(* IEC 61131-3 sources: kns-port-domestic/upstream/kns-pump-station/src/DUTs/Station, 10 files *)

(* ---- E_ControlAct.dut.st ---- *)
// Назначение: действующее управление насосами (04 §4), поле stStationSts.eControlAct.
//             Старшинство в «Автомате»: PowerLost > Restart > DryRunStop > Float > Emergency >
//             LevelPid > Stepped.
// Автор:      kr0nsch
// Версия:     0.1.0
// Документ:   docs/DESIGN.md, раздел 3.1
{attribute 'qualified_only'}
{attribute 'strict'}
TYPE E_ControlAct :
(
    Manual     := 0,   // станция в «Ручном»: запросов нет, только блокировки
    Stepped    := 1,   // ступенчатое регулирование
    LevelPid   := 2,   // ПИД уровня и подключение по нагрузке
    Float      := 3,   // резервное управление по поплавкам (LT101 недостоверен)
    Emergency  := 4,   // аварийно высокий уровень: все доступные насосы
    DryRunStop := 5,   // защита «сухой ход»: запросы сняты
    PowerLost  := 6,   // нет напряжения на вводе
    Restart    := 7    // задержка после старта или восстановления питания, последовательный пуск
) INT;
END_TYPE

(* ---- E_ControlMethod.dut.st ---- *)
// Назначение: выбранный способ регулирования (04 §3.2, 18.2 № 1). Другое значение в retain
//             санитизируется в Stepped.
// Автор:      kr0nsch
// Версия:     0.1.0
// Документ:   docs/DESIGN.md, раздел 3.1
{attribute 'qualified_only'}
{attribute 'strict'}
TYPE E_ControlMethod :
(
    Stepped  := 1,   // ступенчатое по уровням (04 §6)
    LevelPid := 2    // поддержание уровня ПИД LIC101 (04 §7)
) INT;
END_TYPE

(* ---- E_PumpRole.dut.st ---- *)
// Назначение: роль насоса в станции (04 §5.1).
// Автор:      kr0nsch
// Версия:     0.1.0
// Документ:   docs/DESIGN.md, раздел 3.1
{attribute 'qualified_only'}
{attribute 'strict'}
TYPE E_PumpRole :
(
    None    := 0,   // недоступен автоматике (отказ, блокировка, не Auto, нет напряжения)
    Lead    := 1,   // ведущий: запускается первым, в ПИД его частоту регулирует LIC101
    Assist  := 2,   // подпорный: подключается при нехватке производительности
    Standby := 3    // резервный: доступен, не запрошен
) INT;
END_TYPE

(* ---- E_RotationMode.dut.st ---- *)
// Назначение: режим чередования насосов (04 §8.1, 18.2 № 14).
// Автор:      kr0nsch
// Версия:     0.1.0
// Документ:   docs/DESIGN.md, раздел 3.1
{attribute 'qualified_only'}
{attribute 'strict'}
TYPE E_RotationMode :
(
    RunHours := 1,   // по моточасам: меньше RunSeconds, затем меньше Starts, затем меньший номер
    Cyclic   := 2,   // по кругу: следующий после stStationRetain.uiNextLead
    Fixed    := 3    // без чередования: Н1, Н2, Н3
) INT;
END_TYPE

(* ---- E_StationAlarm.dut.st ---- *)
// Назначение: слоты тревог станции KNS1.* (04 §15, 05_alarm_list.csv): индекс массивов
//             FB_StationAlarms и ST_StationCfg.astAlarm; номер тревоги = STN_ALARM_ID_BASE + slot,
//             бит слов wAlm* — slot - 1. Без strict: перечислением индексируются массивы.
// Автор:      kr0nsch
// Версия:     0.1.0
// Документ:   docs/DESIGN.md, раздел 3.1
{attribute 'qualified_only'}
TYPE E_StationAlarm :
(
    EHL    := 1,    // аварийно высокий уровень (Critical)
    DRY    := 2,    // сухой ход станции (High)
    LACK   := 3,    // недостаточно насосов (High)
    NORES  := 4,    // нет резерва (High)
    ATS    := 5,    // АВР выполнен (Medium)
    FLOAT  := 6,    // управление по поплавкам (Medium)
    LDEV   := 7,    // противоречие поплавка и уровнемера (Medium)
    STEP   := 8,    // ступенчатое вместо ПИД (Low)
    NOAUTO := 9,    // станция в «Ручном» дольше 600 с (Low)
    UL1    := 10,   // недогрузка (сухой ход) Н1 (Medium)
    UL2    := 11,   // недогрузка Н2
    UL3    := 12,   // недогрузка Н3
    SIM    := 13    // режим имитации (Low)
) UINT;
END_TYPE

(* ---- E_StationMode.dut.st ---- *)
// Назначение: режим станции (04 §3). Другое значение в retain санитизируется в Manual
//             сравнениями (FB_StationMode, правило L4 контракта plc-process-lib).
// Автор:      kr0nsch
// Версия:     0.1.0
// Документ:   docs/DESIGN.md, раздел 3.1
{attribute 'qualified_only'}
{attribute 'strict'}
TYPE E_StationMode :
(
    Auto   := 1,   // «Автомат»: насосами управляет логика станции
    Manual := 2    // «Ручной»: насосами управляет оператор с HMI, блокировки действуют
) INT;
END_TYPE

(* ---- ST_StationCfg.dut.st ---- *)
// Назначение: уставки станции (GVL_Persist.stStationCfg) — параметры 04 §18.2 № 2–31 с теми же
//             именами и значениями по умолчанию, тревоги KNS1.* и резерв. Значения по умолчанию
//             проходят F_StationCfgCheck. Тип лежит в Persistent Variables и заморожен целиком:
//             новые параметры 1.x — в элементах резерва без переименования.
// Автор:      kr0nsch
// Версия:     0.1.0
// Документ:   docs/DESIGN.md, раздел 3.1
{attribute 'qualified_only'}
TYPE ST_StationCfg :
STRUCT
    // уровни (№ 2–6)
    rLvlStop_m          : REAL := 1.00;
    rLvlStartLead_m     : REAL := 1.60;
    rLvlStopAssist_m    : REAL := 1.40;
    rLvlStartAssist_m   : REAL := 2.40;
    tLvlConfirm         : TIME := T#5S;
    // ступенчатое (№ 7)
    rStepSpeed_pct      : REAL := 100.0;
    // ПИД (№ 8–12)
    rLevelSp_m          : REAL := 1.40;
    rAssistOn_pct       : REAL := 98.0;
    tAssistOn           : TIME := T#30S;
    rAssistOff_pct      : REAL := 75.0;
    tAssistOff          : TIME := T#60S;
    // роли (№ 13–17)
    uiDutyMax           : UINT := 2;
    eRotation           : E_RotationMode := E_RotationMode.RunHours;
    tMaxContRun         : TIME := T#4H;
    tOverlap            : TIME := T#10S;
    tStagger            : TIME := T#5S;
    // питание (№ 18–20)
    tPwrRestart         : TIME := T#10S;
    tSeqStep            : TIME := T#15S;
    tPlcStart           : TIME := T#10S;
    // защиты (№ 21–27)
    tDryRelease         : TIME := T#60S;
    rLdev102On_m        : REAL := 3.50;
    rLdev102Off_m       : REAL := 4.40;
    rLdev103On_m        : REAL := 0.80;
    rLdev103Off_m       : REAL := 0.20;
    tLdev               : TIME := T#30S;
    tLtRecover          : TIME := T#30S;
    // недогрузка (№ 28–30)
    rUnderload_A        : REAL := 12.0;
    rUnderloadSpeed_pct : REAL := 80.0;
    tUnderload          : TIME := T#15S;
    // вентиляция (№ 31)
    tV1Overrun          : TIME := T#10M;
    // тревоги KNS1.* по 05_alarm_list.csv (source = station), индекс — E_StationAlarm. Задержка появления
    // в 05 = tOnDelay + выдержка логики (LDEV — tLdev, UL1…UL3 — tUnderload). Инициализатор — весь
    // массив целиком (правило 3 API 18.3)
    astAlarm            : ARRAY[1..GVL_Const.STN_ALARM_COUNT] OF PL.ST_AlarmCfg := [
        (ePriority := PL.E_AlarmPriority.Critical, tShelveMax := T#0S),   // 1 EHL: откладывать нельзя
        (ePriority := PL.E_AlarmPriority.High),                          // 2 DRY
        (ePriority := PL.E_AlarmPriority.High, tOnDelay := T#10S),       // 3 LACK
        (ePriority := PL.E_AlarmPriority.High, tOnDelay := T#10S),       // 4 NORES
        (ePriority := PL.E_AlarmPriority.Medium),                        // 5 ATS
        (ePriority := PL.E_AlarmPriority.Medium),                        // 6 FLOAT
        (ePriority := PL.E_AlarmPriority.Medium),                        // 7 LDEV
        (ePriority := PL.E_AlarmPriority.Low, tOnDelay := T#10S),        // 8 STEP: без переходных циклов старта
        (ePriority := PL.E_AlarmPriority.Low, tOnDelay := T#10M),        // 9 NOAUTO
        (ePriority := PL.E_AlarmPriority.Medium),                        // 10 UL1
        (ePriority := PL.E_AlarmPriority.Medium),                        // 11 UL2
        (ePriority := PL.E_AlarmPriority.Medium),                        // 12 UL3
        (ePriority := PL.E_AlarmPriority.Low)];                          // 13 SIM
    // резерв: новые параметры 1.x без смены типа; смысл элемента записывается в DESIGN, раздел 3.1
    arReserve           : ARRAY[0..7] OF REAL;
    atReserve           : ARRAY[0..3] OF TIME;
    auiReserve          : ARRAY[0..3] OF UINT;
END_STRUCT
END_TYPE

(* ---- ST_StationCmd.dut.st ---- *)
// Назначение: команды станции (GVL_Station.stStationCmd) — пишут HMI, OPC UA, MQTT. Импульсы и
//             номера обрабатывает и сбрасывает PRG_Station в том же цикле (04 §19.2); результат —
//             stStationSts.eCmdResult и uiCmdSeq.
// Автор:      kr0nsch
// Версия:     0.1.0
// Документ:   docs/DESIGN.md, раздел 3.1
{attribute 'qualified_only'}
TYPE ST_StationCmd :
STRUCT
    xSetAuto      : BOOL;           // импульс: станция в «Автомат» (04 §19.2)
    xSetManual    : BOOL;           // импульс: в «Ручной»; старше xSetAuto
    xSetStepped   : BOOL;           // импульс: способ «ступенчатое»; старше xSetLevelPid
    xSetLevelPid  : BOOL;           // импульс: способ «ПИД уровня»
    xAckAll       : BOOL;           // импульс: квитировать все тревоги станции, LIC101 и устройств
    xResetAll     : BOOL;           // импульс: общий сброс (как HS501)
    xSilence      : BOOL;           // импульс: выключить сирену (как HS502)
    xExportLog    : BOOL;           // импульс: выгрузить журнал в CSV (04 §19.2)
    xRevertCfg    : BOOL;           // импульс: откатить записанные уставки к действующей копии (08 §14, вопрос 2)
    wAckReq       : WORD;           // маска: квитировать тревоги станции, бит slot - 1
    wShelveReq    : WORD;           // маска: отложить на astAlarm[slot].tShelveMax
    wUnshelveReq  : WORD;           // маска: вернуть отложенные
    udiAckId      : UDINT;          // квитировать тревогу по номеру (таблица HMI); 0 — нет; сбрасывается в 0
    udiShelveId   : UDINT;          // отложить тревогу любого источника на её tShelveMax; 0 — нет (08 §14, вопрос 1)
    udiUnshelveId : UDINT;          // вернуть отложенную тревогу по номеру; 0 — нет
END_STRUCT
END_TYPE

(* ---- ST_StationRetain.dut.st ---- *)
// Назначение: энергонезависимое состояние станции (GVL_Persist.stStationRetain): режим, способ
//             регулирования, следующий ведущий для чередования по кругу. Тип лежит в Persistent
//             Variables: не менять (новые данные — в резерве).
// Автор:      kr0nsch
// Версия:     0.1.0
// Документ:   docs/DESIGN.md, раздел 3.1
{attribute 'qualified_only'}
TYPE ST_StationRetain :
STRUCT
    eMode       : E_StationMode := E_StationMode.Manual;      // пустой retain — «Ручной» (04 §3.2)
    eMethod     : E_ControlMethod := E_ControlMethod.Stepped;
    uiNextLead  : UINT := 1;                                  // Cyclic: следующий ведущий
    uiReserve   : UINT;
    audiReserve : ARRAY[0..7] OF UDINT;
END_STRUCT
END_TYPE

(* ---- ST_StationSts.dut.st ---- *)
// Назначение: состояние станции (GVL_Station.stStationSts) для HMI, OPC UA и MQTT: только 16- и
//             32-битные поля, 72 байта (тест StationStsSizeIs72), 04 §19.3.
// Автор:      kr0nsch
// Версия:     0.1.0
// Документ:   docs/DESIGN.md, раздел 3.1
{attribute 'qualified_only'}
TYPE ST_StationSts :
STRUCT
    eMode             : E_StationMode;
    eMethod           : E_ControlMethod;
    eControlAct       : E_ControlAct;
    eNe107            : PL.E_Ne107Status;   // F — LACK; S — FLOAT, STEP, LDEV, NORES; C — «Ручной», имитация,
                                            // wCfgErr; M — ТО насоса
    wState            : WORD;               // биты STN_ST_*
    wCfgErr           : WORD;               // биты STN_CFG_*
    aeRole            : ARRAY[1..3] OF E_PumpRole;
    uiPumpsRequired   : UINT;
    uiPumpsRunning    : UINT;
    uiPumpsAvailable  : UINT;
    uiLeadPump        : UINT;               // 0 — нет
    uiSeqRemain_s     : UINT;
    eCmdResult        : PL.E_CmdResult;     // результат последней команды станции
    uiCmdSeq          : UINT;               // +1 на каждую обработанную команду
    wAlmActive        : WORD;               // тревоги станции, бит slot - 1
    wAlmUnack         : WORD;
    wAlmShelved       : WORD;               // дополнение: Shelved, SuppressedByDesign, OutOfService
    ePrioUnack        : PL.E_AlarmPriority; // высший неквитированный по всем источникам (баннер)
    auiUnack          : ARRAY[1..4] OF UINT;// неквитированных Low…Critical
    eLogExport        : E_LogExportState;   // дополнение: состояние выгрузки CSV
    wReserve          : WORD;               // выравнивание: дальше 32-битные поля
    rLevel_m          : REAL;               // уровень, по которому работает станция
    rLevelSp_m        : REAL;               // действующее задание уровня
    rSpeedSp_pct      : REAL;               // общее задание частоты насосам
    udiEventSeq       : UDINT;              // номер последней записи журнала
    udiLogOverwritten : UDINT;              // затёрто записей журнала
END_STRUCT
END_TYPE
